// TIA Portal V21 export
FUNCTION_BLOCK "FB_AnaTimerCaller"   // FB19, SCL
TITLE = Analyzer: FB with a timer called inside IF
{ S7_Optimized_Access := 'TRUE' }
// Rule C26m (caller): FB_AnaTimerInner contains a timer and is called only while Enable is TRUE
// stored: MemoryReserve 100, SetENOAutomatically false
   VAR_INPUT
      Enable : Bool;   // Enable
      Start : Bool;   // Start of the inner timer
   END_VAR
   VAR_OUTPUT
      Done : Bool;   // Output of the inner timer
   END_VAR
   VAR
      Inner { S7_SetPoint := 'True'} : "FB_AnaTimerInner";   // FB that contains a timer
   END_VAR
BEGIN

       IF #Enable THEN
           #Inner(Start := #Start);
       END_IF;
       #Done := #Inner.Done;
END_FUNCTION_BLOCK
